FUNCTION_BLOCK TransportToClient (* Composite Function Block Type *)
  (* Standard: 61499-2 *)
  (* Version 0.0, 7/2/2026, template *)
  PACKAGE Main;
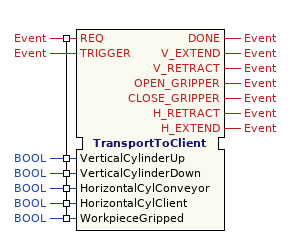
  EVENT_INPUT
    REQ WITH VerticalCylinderUp, VerticalCylinderDown, HorizontalCylConveyor, HorizontalCylClient, WorkpieceGripped; (* Normal Execution Request *)
    TRIGGER;
  END_EVENT
  EVENT_OUTPUT
    DONE;
    V_EXTEND;
    V_RETRACT;
    OPEN_GRIPPER;
    CLOSE_GRIPPER;
    H_RETRACT;
    H_EXTEND;
  END_EVENT
  VAR_INPUT
    VerticalCylinderUp : BOOL; (* Input event qualifier *)
    VerticalCylinderDown : BOOL;
    HorizontalCylConveyor : BOOL;
    HorizontalCylClient : BOOL;
    WorkpieceGripped : BOOL;
  END_VAR
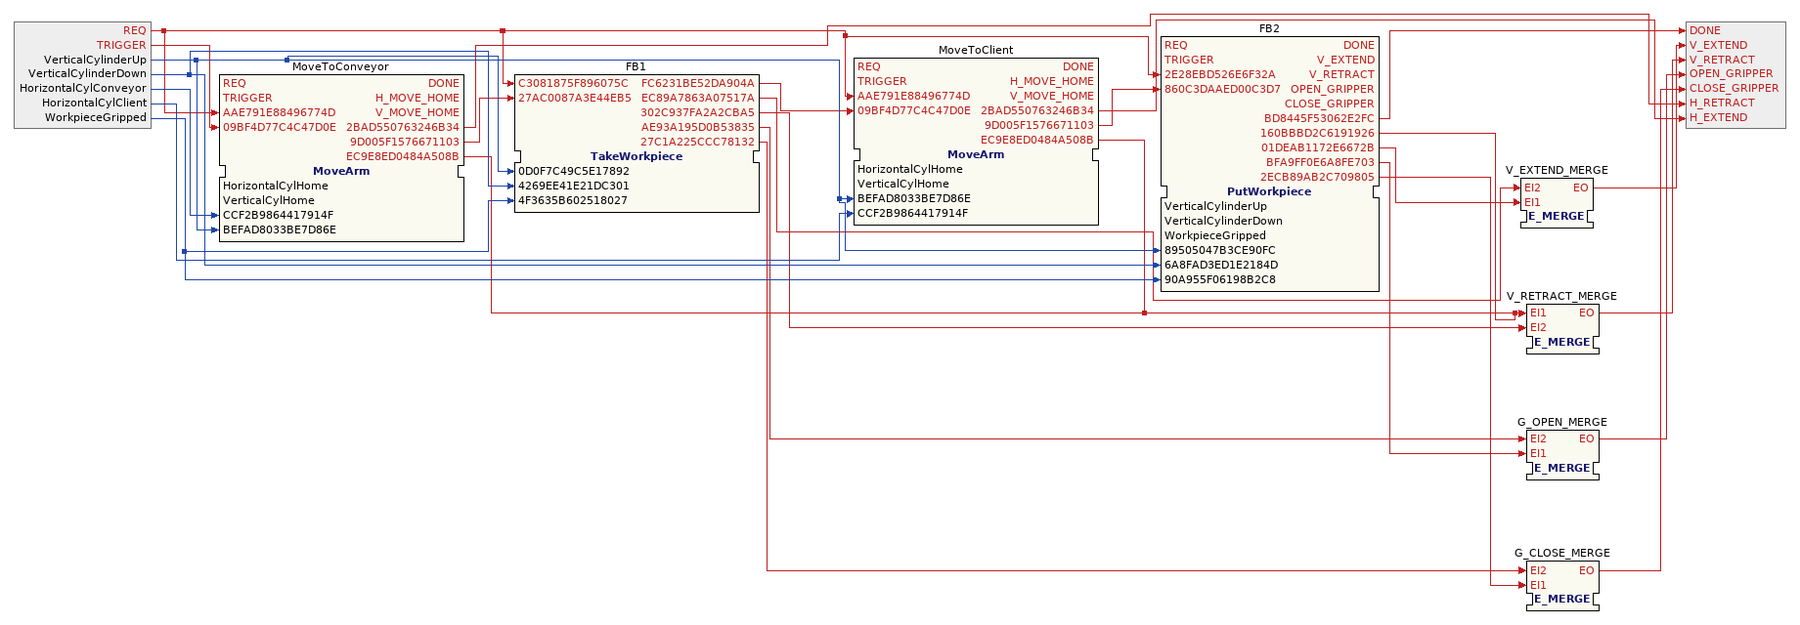
  FBS
    MoveToConveyor : MoveArm;
    FB1 : TakeWorkpiece;
    MoveToClient : MoveArm;
    FB2 : PutWorkpiece;
    V_EXTEND_MERGE : E_MERGE;
    V_RETRACT_MERGE : E_MERGE;
    G_OPEN_MERGE : E_MERGE;
    G_CLOSE_MERGE : E_MERGE;
  END_FBS
  EVENT_CONNECTIONS
    FB2.BD8445F53062E2FC TO DONE;
    V_EXTEND_MERGE.EO TO V_EXTEND;
    V_RETRACT_MERGE.EO TO V_RETRACT;
    G_OPEN_MERGE.EO TO OPEN_GRIPPER;
    G_CLOSE_MERGE.EO TO CLOSE_GRIPPER;
    MoveToClient.2BAD550763246B34 TO H_EXTEND;
    MoveToConveyor.2BAD550763246B34 TO H_RETRACT;
    REQ TO MoveToConveyor.AAE791E88496774D;
    REQ TO FB1.C3081875F896075C;
    REQ TO MoveToClient.AAE791E88496774D;
    REQ TO FB2.2E28EBD526E6F32A;
    MoveToClient.9D005F1576671103 TO FB2.860C3DAAED00C3D7;
    FB1.FC6231BE52DA904A TO MoveToClient.09BF4D77C4C47D0E;
    MoveToConveyor.9D005F1576671103 TO FB1.27AC0087A3E44EB5;
    TRIGGER TO MoveToConveyor.09BF4D77C4C47D0E;
    MoveToConveyor.EC9E8ED0484A508B TO V_RETRACT_MERGE.EI1;
    FB1.EC89A7863A07517A TO V_EXTEND_MERGE.EI2;
    FB1.302C937FA2A2CBA5 TO V_RETRACT_MERGE.EI2;
    FB1.AE93A195D0B53835 TO G_OPEN_MERGE.EI2;
    FB1.27C1A225CCC78132 TO G_CLOSE_MERGE.EI2;
    MoveToClient.EC9E8ED0484A508B TO V_RETRACT_MERGE.EI1;
    FB2.160BBBD2C6191926 TO V_RETRACT_MERGE.EI1;
    FB2.01DEAB1172E6672B TO V_EXTEND_MERGE.EI1;
    FB2.BFA9FF0E6A8FE703 TO G_OPEN_MERGE.EI1;
    FB2.2ECB89AB2C709805 TO G_CLOSE_MERGE.EI1;
  END_CONNECTIONS
  DATA_CONNECTIONS
    HorizontalCylConveyor TO MoveToConveyor.CCF2B9864417914F;
    VerticalCylinderUp TO MoveToConveyor.BEFAD8033BE7D86E;
    VerticalCylinderUp TO FB1.0D0F7C49C5E17892;
    VerticalCylinderUp TO MoveToClient.BEFAD8033BE7D86E;
    VerticalCylinderUp TO FB2.89505047B3CE90FC;
    VerticalCylinderDown TO FB1.4269EE41E21DC301;
    VerticalCylinderDown TO FB2.6A8FAD3ED1E2184D;
    HorizontalCylClient TO MoveToClient.CCF2B9864417914F;
    WorkpieceGripped TO FB1.4F3635B602518027;
    WorkpieceGripped TO FB2.90A955F06198B2C8;
  END_CONNECTIONS
END_FUNCTION_BLOCK
